(* Simple Agitated Mixing Tank with Heater Coil *)

PROGRAM main
  VAR
    InletValve1 AT %QX0.1 : BOOL; (* Output Device for Material A Intake *)
    InletValve2 AT %QX0.2 : BOOL; (* Output Device for Material B Intake *)
    OutletValve AT %QX0.6 : BOOL;
    Start AT %IX0.1 : BOOL; (* Simple Push Button Input *)
    Stop AT %IX0.2 : BOOL; (* Simple Push Button Input *)
    CycleOn AT %QX0.3 : BOOL;
    LevelSensor1 AT %IX0.4 : BOOL; (* Upper Level Sensor *)
    LevelSensor2 AT %IX0.5 : BOOL;
    LowLevelSensor AT %IX0.6 : BOOL; (* Tank Empty Sensor *)
    AgitatorMotor AT %QX0.4 : BOOL; (* Actuator for Mixing Materials *)
    Heater AT %QX0.5 : BOOL;
    Flag AT %MX0.1 : BOOL;
    TemperatureSensor AT %IW1 : INT;
    TP0 : TP;
  END_VAR

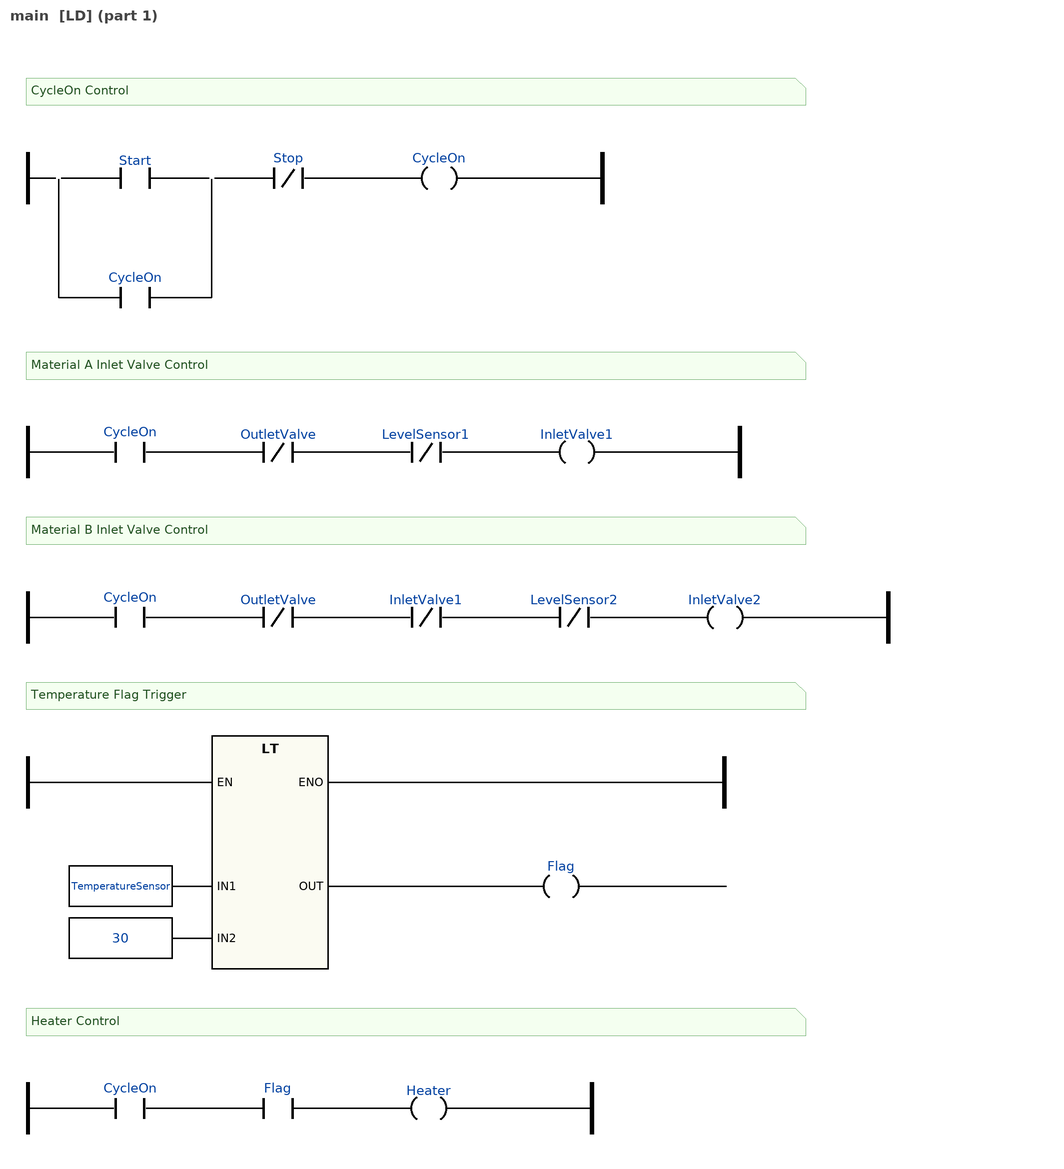
(* LD diagram, written out as Structured Text *)
(* CycleOn Control *)
CycleOn := (Start OR CycleOn) AND NOT Stop;
(* Material A Inlet Valve Control *)
InletValve1 := CycleOn AND NOT OutletValve AND NOT LevelSensor1;
(* Material B Inlet Valve Control *)
InletValve2 := CycleOn AND NOT OutletValve AND NOT InletValve1 AND NOT LevelSensor2;
(* Temperature Flag Trigger *)
Flag := TemperatureSensor < 30;
(* Heater Control *)
Heater := CycleOn AND Flag;
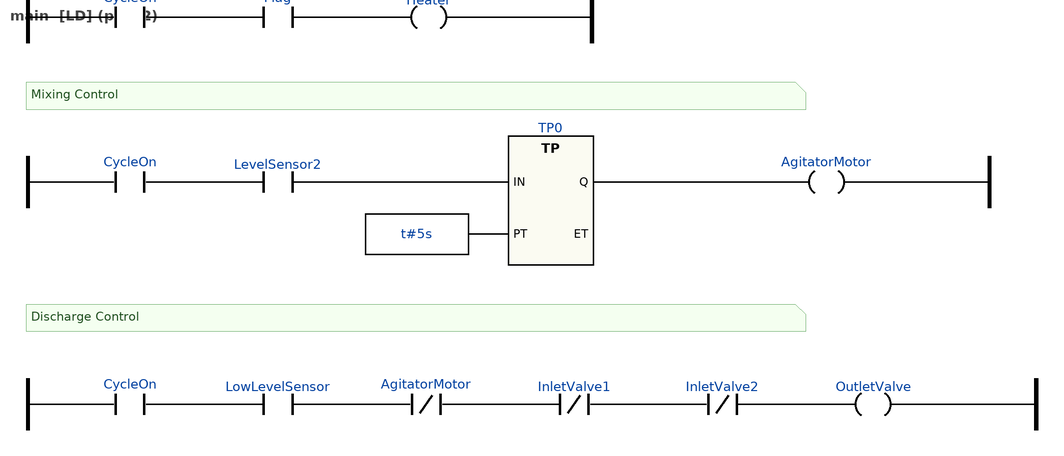
(* Mixing Control *)
TP0(IN := CycleOn AND LevelSensor2, PT := t#5s);
AgitatorMotor := TP0.Q;
(* Discharge Control *)
OutletValve := CycleOn AND LowLevelSensor AND NOT AgitatorMotor AND NOT InletValve1 AND NOT InletValve2;
END_PROGRAM
